// TIA Portal V20 export
// export: Created 2026-10-20T18:54:44.0018117Z, ExportSetting None, DisplayName Totally Integrated Automation Portal, DisplayVersion V20 Update 6, DisplayName TIA Portal Openness, DisplayVersion V20 Update 6, DisplayName TIA Portal Version Control Interface, DisplayVersion V20 Update 6, DisplayName SINAMICS Startdrive Advanced, DisplayVersion V20 SP1, DisplayName SINAMICS Startdrive G130, G150, S120, S150, SINAMICS MV, G220, S200, S210, DisplayVersion V20 SP1, DisplayName SINAMICS Startdrive G110M, G120, G120C, G120D, G120P, G115D, DisplayVersion V20 SP1, DisplayName STEP 7 Professional, DisplayVersion V20 Update 6, DisplayName STEP 7 Safety, DisplayVersion V20 Update 2, DisplayName WinCC Basic/Comfort/Advanced, DisplayVersion V20 Update 6, DisplayName WinCC Unified, DisplayVersion V20 Update 6
VAR_GLOBAL   // PLC tag table "IO_VFDs_1"
   VTD1_ControlWord AT %QW40 : Word;
   VTD1_MainSetpoint AT %QW42 : Word;
   VTD1_StatusWord AT %IW44 : Word;
   VTD1_ActualSpeed AT %IW46 : Word;
   VTD1_ActualCurrent AT %IW48 : Word;
   C1101_ControlWord AT %QW50 : Word;
   C1101_MainSetpoint AT %QW52 : Word;
   C1101_StatusWord AT %IW2018 : Word;
   C1101_ActualSpeed AT %IW2020 : Word;
   C1101_ActualCurrent AT %IW2022 : Word;
   C1102_ControlWord AT %QW54 : Word;
   C1102_MainSetpoint AT %QW56 : Word;
   C1102_StatusWord AT %IW2030 : Word;
   C1102_ActualSpeed AT %IW2032 : Word;
   C1102_ActualCurrent AT %IW2034 : Word;
   C1103_ControlWord AT %QW58 : Word;
   C1103_MainSetpoint AT %QW60 : Word;
   C1103_StatusWord AT %IW2042 : Word;
   C1103_ActualSpeed AT %IW2044 : Word;
   C1103_ActualCurrent AT %IW2046 : Word;
   C1104_ControlWord AT %QW62 : Word;
   C1104_MainSetpoint AT %QW64 : Word;
   C1104_StatusWord AT %IW2054 : Word;
   C1104_ActualSpeed AT %IW2056 : Word;
   C1104_ActualCurrent AT %IW2058 : Word;
   C1105_ControlWord AT %QW66 : Word;
   C1105_MainSetpoint AT %QW68 : Word;
   C1105_StatusWord AT %IW2066 : Word;
   C1105_ActualSpeed AT %IW2068 : Word;
   C1105_ActualCurrent AT %IW2070 : Word;
   C1106_ControlWord AT %QW70 : Word;
   C1106_MainSetpoint AT %QW72 : Word;
   C1106_StatusWord AT %IW2078 : Word;
   C1106_ActualSpeed AT %IW2080 : Word;
   C1106_ActualCurrent AT %IW2082 : Word;
   C1107_ControlWord AT %QW186 : Word;
   C1107_MainSetpoint AT %QW188 : Word;
   C1107_StatusWord AT %IW2198 : Word;
   C1107_ActualSpeed AT %IW2200 : Word;
   C1107_ActualCurrent AT %IW2202 : Word;
   CVTD1_ControlWord AT %QW46 : Word;
   CVTD1_MainSetpoint AT %QW48 : Word;
   CVTD1_StatusWord AT %IW2006 : Word;
   CVTD1_ActualSpeed AT %IW2008 : Word;
   CVTD1_ActualCurrent AT %IW2010 : Word;
   C1108_ControlWord AT %QW74 : Word;
   C1108_MainSetpoint AT %QW76 : Word;
   C1108_StatusWord AT %IW2090 : Word;
   C1108_ActualSpeed AT %IW2092 : Word;
   C1108_ActualCurrent AT %IW2094 : Word;
   C1201_ActualCurrent AT %IW2106 : Word;
   C1201_ActualSpeed AT %IW2104 : Word;
   C1201_ControlWord AT %QW78 : Word;
   C1201_MainSetpoint AT %QW80 : Word;
   C1201_StatusWord AT %IW2102 : Word;
   C1202_ActualCurrent AT %IW2118 : Word;
   C1202_ActualSpeed AT %IW2116 : Word;
   C1202_ControlWord AT %QW82 : Word;
   C1202_MainSetpoint AT %QW84 : Word;
   C1202_StatusWord AT %IW2114 : Word;
   C1203_ActualCurrent AT %IW2130 : Word;
   C1203_ActualSpeed AT %IW2128 : Word;
   C1203_ControlWord AT %QW86 : Word;
   C1203_MainSetpoint AT %QW88 : Word;
   C1203_StatusWord AT %IW2126 : Word;
   C1204_ActualCurrent AT %IW2142 : Word;
   C1204_ActualSpeed AT %IW2140 : Word;
   C1204_ControlWord AT %QW90 : Word;
   C1204_MainSetpoint AT %QW92 : Word;
   C1204_StatusWord AT %IW2138 : Word;
   C1205_ActualCurrent AT %IW2154 : Word;
   C1205_ActualSpeed AT %IW2152 : Word;
   C1205_ControlWord AT %QW94 : Word;
   C1205_MainSetpoint AT %QW96 : Word;
   C1205_StatusWord AT %IW2150 : Word;
   C1206_ActualCurrent AT %IW2166 : Word;
   C1206_ActualSpeed AT %IW2164 : Word;
   C1206_ControlWord AT %QW174 : Word;
   C1206_MainSetpoint AT %QW176 : Word;
   C1206_StatusWord AT %IW2162 : Word;
   C1207_ActualCurrent AT %IW2178 : Word;
   C1207_ActualSpeed AT %IW2176 : Word;
   C1207_ControlWord AT %QW178 : Word;
   C1207_MainSetpoint AT %QW180 : Word;
   C1207_StatusWord AT %IW2174 : Word;
   C1208_ActualCurrent AT %IW2190 : Word;
   C1208_ActualSpeed AT %IW2188 : Word;
   C1208_ControlWord AT %QW182 : Word;
   C1208_MainSetpoint AT %QW184 : Word;
   C1208_StatusWord AT %IW2186 : Word;
   C1201_ActualTorque AT %IW2108 : Word;
   C1101_ActualTorque AT %IW2024 : Word;
   C1107_ActualTorque AT %IW2204 : Word;
   VTD1_ActualTorque AT %IW50 : Word;
   C1108_ActualTorque AT %IW2096 : Word;
   C1103_ActualTorque AT %IW2048 : Word;
   C1105_ActualTorque AT %IW2072 : Word;
   C1102_ActualTorque AT %IW2036 : Word;
   C1203_ActualTorque AT %IW2132 : Word;
   C1104_ActualTorque AT %IW2060 : Word;
   C1207_ActualTorque AT %IW2180 : Word;
   C1204_ActualTorque AT %IW2144 : Word;
   C1202_ActualTorque AT %IW2120 : Word;
   C1206_ActualTorque AT %IW2168 : Word;
   C1106_ActualTorque AT %IW2084 : Word;
   C1208_ActualTorque AT %IW2192 : Word;
   CVTD1_ActualTorque AT %IW2012 : Word;
   C1205_ActualTorque AT %IW2156 : Word;
   VTD1_AccFactor AT %QW1513 : Word;
END_VAR
